(* IEC 61131-3 sources: plc-vscode/tests/st/test-ready/rusty/tests/lit/single/auto_pointers, 3 files *)

(* ---- var_in_out_array_of_array_scalar.st ---- *)
// RUN: (%COMPILE %s && %RUN) | %CHECK %s
// XFAIL: *
// failing because of #1508
FUNCTION foo
VAR_IN_OUT
    in : ARRAY[0..1] OF ARRAY[0..1] OF INT;
END_VAR
    in[0][0] := 1;
    in[0][1] := 2;
    in[1][0] := 3;
    in[1][1] := 4;
END_FUNCTION

FUNCTION main
VAR
    arr: ARRAY[0..1] OF ARRAY[0..1] OF INT;
END_VAR
    foo(arr);
    // CHECK: 1 2 3 4
    printf('%d %d %d %d$N', arr[0][0], arr[0][1], arr[1][0], arr[1][1]);
END_FUNCTION

(* ---- var_in_out_array_of_string.st ---- *)
// RUN: (%COMPILE %s && %RUN) | %CHECK %s
FUNCTION foo
VAR_IN_OUT
    in_out : ARRAY[0..3] OF STRING;
END_VAR
VAR_INPUT {ref}
    in: ARRAY[0..3] OF STRING;
END_VAR
    in_out[0] := 'YOU';
    in_out[1] := 'SHALL';
    in[2] := 'NOT';
    in[3] := 'SEGFAULT';
END_FUNCTION

FUNCTION main
VAR
    arr: ARRAY[0..3] OF STRING;
END_VAR
    foo(arr, arr);
    // CHECK: YOU SHALL NOT SEGFAULT
    printf('%s %s %s %s$N', REF(arr[0]), REF(arr[1]), REF(arr[2]), REF(arr[3]));
END_FUNCTION

(* ---- var_in_out_strings_with_different_lengths.st ---- *)
// RUN: (%COMPILE %s && %RUN) | %CHECK %s
FUNCTION foo
VAR_IN_OUT
    str80_io : STRING;
    str10_io : STRING[10];
END_VAR
    str80_io := 'hello';
    str10_io := 'ralph';
END_FUNCTION

FUNCTION main
VAR
    str80 : STRING;
    str10 : STRING[10];
END_VAR
    foo(str80, str10);
    // CHECK: ralph hello
    printf('%s %s$N', REF(str10), REF(str80));
END_FUNCTION
